PROGRAM MAIN
VAR
	//instantiation of the test case function blocks
	fbT1	: FB_TestSum;   //Test case for the FB_Sum function block from the library
	fbT2	: FB_TestDiff;  //Test case for the FB_Diff function block from the library
	fbT3	: FB_TestProd;  //Test case for the FB_Prod function block from the library
	fbT4	: FB_TestDiv;   //Test case for the FB_Div function block from the library
END_VAR

//To have the source code for a library’s unit tests directly within the same solution, it is advisable to enable the option “Allow the project to be referenced as a library” in the library project. This option makes it possible to run the tests at any time without having to install the library on the system. It is therefore particularly useful for use in CI/CD pipelines, as the command to install the libraries does not need to be executed.

// Calling the TestController (which is located in the library and acts as the interface to the clients) 
Tc3_PlcTestFramework.F_CallTestController();

END_PROGRAM

(* stored: Version 1.1.0.1, ProductVersion 3.1.4026.21
   POU MAIN: Id {359411d8-4113-43aa-ae2e-7e41eef1cef1}, SpecialFunc None *)
